// TIA Portal V21 export
// export: Created 2026-11-08T21:46:52.2299481Z, ExportSetting WithDefaults, DisplayName Totally Integrated Automation Portal, DisplayVersion V21 Update 3, DisplayName STEP 7 Professional, DisplayVersion V21 Update 3, DisplayName STEP 7 Safety, DisplayVersion V21, DisplayName Tech WebApplication, DisplayVersion V21, DisplayName WinCC Basic/Comfort/Advanced, DisplayVersion V21 Update 3, DisplayName WinCC Unified, DisplayVersion V21 Update 3
DATA_BLOCK "DB_Khp"   // DB6
{ S7_Optimized_Access := 'TRUE' }
VERSION : 0.1
// stored: AutoNumber true, DBAccessibleFromOPCUA true, DBAccessibleFromWebserver true, IsOnlyStoredInLoadMemory false, IsRetainMemResEnabled false, IsWriteProtectedInAS false, MemoryReserve 100
   VAR
      "a" : Int := 7;
      "b" : Real := 1.5;
      s : Struct
         x : Bool;
         y : Array[0..2] of DInt;
      END_STRUCT;
      "m" { S7_SetPoint := 'True'} : "UDT_Motor";
   END_VAR
BEGIN
   s.y[1] := 11;
END_DATA_BLOCK
